(* IEC 61131-3 sources: model-first-plc-agent-ai/results/T1-W-14, 2 files *)

(* ---- a1_code.st ---- *)
FUNCTION_BLOCK TransferRuntime
VAR_INPUT
    initialize : BOOL;
    sensor_a : BOOL;
    sensor_b : BOOL;
END_VAR
VAR_OUTPUT
    conveyor : BOOL;
END_VAR
VAR
    command_latch : RS;
END_VAR

(* Initialize G1 to x0: conveyor stopped. *)
IF initialize THEN
    command_latch(S := FALSE, R1 := TRUE);
END_IF;

(* Reset dominance implements both GRAFCET transitions:
   x0 -> x1 when sensor_a AND NOT sensor_b;
   x1 -> x0 when sensor_b. *)
command_latch(
    S := sensor_a AND NOT sensor_b,
    R1 := sensor_b
);

conveyor := command_latch.Q1;

END_FUNCTION_BLOCK

PROGRAM Main
VAR
    SensorA AT %IX100.0 : BOOL;
    SensorB AT %IX100.1 : BOOL;
    Conveyor AT %QX100.0 : BOOL;
END_VAR
VAR
    runtime_logic : TransferRuntime;
    first_scan : BOOL := TRUE;
END_VAR

runtime_logic(
    initialize := first_scan,
    sensor_a := SensorA,
    sensor_b := SensorB
);

Conveyor := runtime_logic.conveyor;
first_scan := FALSE;

END_PROGRAM

(* ---- a2_code.st ---- *)
FUNCTION_BLOCK FB_ConveyorControl
VAR_INPUT
    sensor_a : BOOL;
    sensor_b : BOOL;
END_VAR
VAR_OUTPUT
    conveyor : BOOL;
END_VAR
VAR
    command_latch : RS;
END_VAR

command_latch(S := sensor_a, R1 := sensor_b);
conveyor := command_latch.Q1;

END_FUNCTION_BLOCK

PROGRAM Main
VAR
    sensor_a AT %IX100.0 : BOOL;
    sensor_b AT %IX100.1 : BOOL;
    conveyor AT %QX100.0 : BOOL;
END_VAR
VAR
    controller : FB_ConveyorControl;
END_VAR

controller(sensor_a := sensor_a, sensor_b := sensor_b);
conveyor := controller.conveyor;

END_PROGRAM
